// TIA Portal V20 export
// export: Created 2026-10-30T22:15:00.2103700Z, ExportSetting WithDefaults
ORGANIZATION_BLOCK "Jumps"   // OB1, LAD, ProgramCycle
{ S7_Optimized_Access := 'TRUE' }
VERSION : 0.1
// stored: AutoNumber true, IsIECCheckEnabled true, SetENOAutomatically false
   VAR_INPUT
      Initial_Call : Bool;
   END_VAR
   VAR_TEMP
      valA : DInt;
      valB : DInt;
      valC : DInt;
      result : DInt;
      selector : USInt;
      caseA : USInt;
      caseB : USInt;
      done : Bool;
   END_VAR
BEGIN

REGION Network 1: Switch
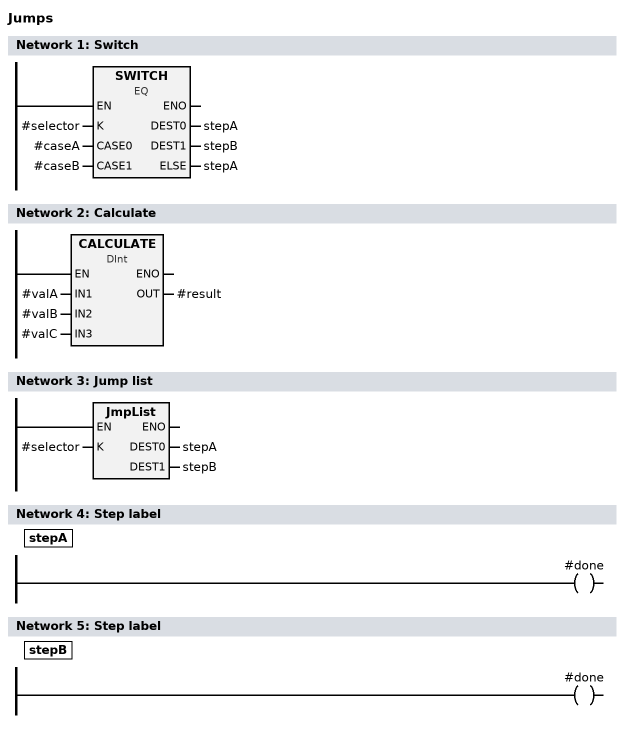
   // no SCL statement known for Switch: written as a call
   Switch(k := #selector, case0 := #caseA, case1 := #caseB, dest0 => stepA, dest1 => stepB, "else" => stepA);
END_REGION

REGION Network 2: Calculate
   RUNG wire#powerrail
      { S7_Templates := "SrcType := DInt"; S7_Expression := "(IN1 + IN2) * (IN1 - IN2)" } Calculate(in1 := #valA, in2 := #valB, in3 := #valC, out => #result)
   END_RUNG
   // the same network as SCL:
   #result := (#valA + #valB) * (#valA - #valB);
END_REGION

REGION Network 3: Jump list
   // no SCL statement known for JmpList: written as a call
   JmpList(k := #selector, dest0 => stepA, dest1 => stepB);
END_REGION

REGION Network 4: Step label
   Label( stepA )
   RUNG wire#powerrail
      Coil( #done )
   END_RUNG
   // the same network as SCL:
   stepA:
   #done := TRUE;
END_REGION

REGION Network 5: Step label
   Label( stepB )
   RUNG wire#powerrail
      Coil( #done )
   END_RUNG
   // the same network as SCL:
   stepB:
   #done := TRUE;
END_REGION
END_ORGANIZATION_BLOCK
